    rq_activate_all_grippers(True)
    # end: URCap Program Node
  end
  $ 63 "zero_ftsensor()"
  zero_ftsensor()
  $ 64 "EXTT"
  $ 65 "Set GRP_3F_Enable=Off"
  set_standard_digital_out(4, False)
  $ 66 "Set BarcodeTrigger=Off"
  set_standard_digital_out(6, False)
  $ 67 "Set GRP_3F_Decap=Off"
  set_standard_digital_out(3, False)
  $ 68 "Set GRP_3F_Cap=Off"
  set_standard_digital_out(2, False)
  $ 69 "Set GRP_3F_Open=Off"
  set_standard_digital_out(5, False)
  $ 70 "PSE_T≔get_tool_free_pose(dir=[0,0,0.150], move_in_base_frame=True)"
  global PSE_T=get_tool_free_pose(dir=[0,0,0.150], move_in_base_frame=True)
  $ 71 "If is_reachable(Base_const, [PSE_T])"
  if (is_reachable(p[0.0,0.0,0.0,0.0,0.0,0.0], [PSE_T])):
    $ 72 "MoveL"
    $ 73 "PSE_T" "breakAfter"
    movel(PSE_T, a=1.2, v=0.15)
  end
  $ 74 "powder dispensing variable init"
  $ 75 "Start_thread≔ False "
  global Start_thread=  False
  $ 76 "vib_thread≔ False "
  global vib_thread=  False
  $ 77 "kp≔0.001"
  global kp=0.001
  $ 78 "ki≔0.00006"
  global ki=0.00006
  $ 79 "kd≔0.015"
  global kd=0.015
  $ 80 "dt≔0.03"
  global dt=0.03
  $ 81 "Integral_error≔0"
  global Integral_error=0
  $ 82 "current_error≔0"
  global current_error=0
  $ 83 "previous_error≔0"
  global previous_error=0
  $ 84 "tilt_increment≔0"
  global tilt_increment=0
  $ 85 "tilt_angle≔0"
  global tilt_angle=0
  $ 86 "diff≔0"
  global diff=0
  $ 87 "current_pose≔get_actual_tcp_pose()"
  global current_pose= get_actual_tcp_pose ()
  $ 88 "Relative_trans≔p[0, 0, -0.035, 0, 0, 0]"
  global Relative_trans=p[0, 0, -0.035, 0, 0, 0]
  $ 89 "ContA_plc_offst≔p[-0.00205, 0.02547, 0.03730, -0.03, -2.183, 6.165]"
  global ContA_plc_offst=p[-0.00205, 0.02547, 0.03730, -0.03, -2.183, 6.165]
  $ 90 "PowA_50_offset≔p[0.21808, -0.19943, 0.06584, 0, 0, 0]"
  global PowA_50_offset=p[0.21808, -0.19943, 0.06584, 0, 0, 0]
  $ 92 "tilt_init_reference()"
  tilt_init_reference()
  $ 93 "switch_spat_M≔ True "
  global switch_spat_M=  True
  $ 94 "switch_spat_S≔ True "
  global switch_spat_S=  True
  $ 95 "switch_spat_F_M≔ True "
  global switch_spat_F_M=  True
  $ 96 "switch_spat_F_S≔ True "
  global switch_spat_F_S=  True
  $ 97 "last_scale≔0"
  global last_scale=0
  $ 98 "W_EMPTY≔51.3"
  global W_EMPTY=51.3
  $ 99 "w_dosed_total≔0"
  global w_dosed_total=0
  $ 794 "Thread_1"
  thread Thread_1():
    while (True):
      $ 795 "If Start_thread≟ True "
      if (Start_thread ==   True  ):
        $ 796 "weight_value≔get_weight()"
        global weight_value=get_weight()
        $ 797 "Wait: 0.1"
        sleep(0.1)
        $ 798 "sync()"
        sync()
      end
      $ 799 "sync()"
      sync()
    end
  end
  threadId_Thread_1 = run Thread_1()
  $ 800 "Thread_2"
  thread Thread_2():
    while (True):
      $ 801 "Loop vib_thread≟ True "
      thread Thread_while_801():
        while (True):
          $ 802 "diff≔target_weight-weight_value"
          global diff=target_weight-weight_value
          $ 803 "If diff>0.02 and spatula≠'spatula_flat_S'"
          global thread_flag_803=0
          thread Thread_if_803():
            $ 805 "Set AO[0]=4.0"
            set_standard_analog_out(0, 0.4)
            thread_flag_803 = 1
          end
          if (diff>0.02  and  spatula != "spatula_flat_S"):
            global thread_handler_803=run Thread_if_803()
            while (thread_flag_803 == 0):
              if not(diff>0.02  and  spatula != "spatula_flat_S"):
                kill thread_handler_803
                thread_flag_803 = 2
              else:
                sync()
              end
            end
          else:
            thread_flag_803 = 2
          end
          if (thread_flag_803 == 2):
            $ 806 "ElseIf diff>0.02 and spatula≟'spatula_flat_S'"
            if (diff>0.02 and spatula == "spatula_flat_S"):
              $ 807 "vibration_3()"
              vibration_3()
            else:
              $ 808 "ElseIf diff≤0.03"
              global thread_flag_808=0
              thread Thread_if_808():
                $ 809 "vibration_2()"
                vibration_2()
                thread_flag_808 = 1
              end
              if (diff <= 0.03):
                global thread_handler_808=run Thread_if_808()
                while (thread_flag_808 == 0):
                  if not(diff <= 0.03):
                    kill thread_handler_808
                    thread_flag_808 = 2
                  else:
                    sync()
                  end
                end
              else:
                thread_flag_808 = 2
              end
              if (thread_flag_808 == 2):
                $ 814 "Else" "noBreak"
                $ 815 "Set AO[0]=0.0"
                set_standard_analog_out(0, 0.0)
              end
            end
          end
        end
      end
      if (vib_thread ==   True  ):
        global thread_handler_801=run Thread_while_801()
        while (vib_thread ==   True  ):
          sync()
        end
        kill thread_handler_801
      end
      $ 816 "sync()"
      sync()
    end
  end
  threadId_Thread_2 = run Thread_2()
  while (True):
    $ 100 "Robot Program"
    $ 101 "MAIN"
    $ 102 "command_manager(external_control='uGO', cond_suspend=(ITM_Manipulated and AMR_AtTarget and AMR_Charging and AMR_Battery<40), cond_unsuspend=(AMR_Battery≟60))"
    command_manager(external_control="uGO", cond_suspend=(ITM_Manipulated  and  AMR_AtTarget  and  AMR_Charging  and  AMR_Battery<40), cond_unsuspend=(AMR_Battery == 60))
    $ 103 "log_state(STATE_Info)"
    log_state(STATE_Info)
    $ 104 "Switch STATE"
    switch_1 = STATE
    $ 105 "Case 1"
    if (1 == switch_1):
      $ 106 "Stopping"
      $ 107 "STATE_Info≔'Stopping'"
      global STATE_Info="Stopping"
      $ 108 "end_freedrive_mode()"
      end_freedrive_mode()
      $ 109 "Set"
      set_tcp(p[0.0,0.0,0.161,3.1415,0.0,0.0])
      $ 110 "PSE_T≔get_tool_free_pose(dir=[0,0,0.150], move_in_base_frame=True)"
      global PSE_T=get_tool_free_pose(dir=[0,0,0.150], move_in_base_frame=True)
      $ 111 "If is_reachable(Base_const, [PSE_T])"
      if (is_reachable(p[0.0,0.0,0.0,0.0,0.0,0.0], [PSE_T])):
        $ 112 "MoveL"
        $ 113 "PSE_T" "breakAfter"
        movel(PSE_T, a=1.2, v=0.15)
      end
      $ 114 "do_transition(keep_rxry=OBJ_Picked, r=0)"
      do_transition(keep_rxry=OBJ_Picked, r=0)
      $ 123 "Call Sub_AMR_MiR_V3"
      Sub_AMR_MiR_V3()
      $ 124 "If stopping() and AMR_Done"
      if (stopping()  and  AMR_Done):
        $ 125 "STATE≔2"
        global STATE=2
        $ 126 "ugo_update_outputs()"
        ugo_update_outputs()
      end
    elif (2 == switch_1):
      $ 127 "Case 2"
      $ 128 "Stopped"
      $ 129 "STATE_Info≔'Stopped'"
      global STATE_Info="Stopped"
      $ 130 "Call Sub_AMR_MiR_V3"
      Sub_AMR_MiR_V3()
      $ 131 "If CMD_Reset  or PB_Start"
      if (CMD_Reset   or  get_standard_digital_in(0)):
        $ 132 "STATE≔3"
        global STATE=3
        $ 133 "ugo_update_outputs()"
        ugo_update_outputs()
      end
    elif (3 == switch_1):
      $ 134 "Case 3"
      $ 135 " Resetting"
      $ 136 "STATE_Info≔'Resetting'"
      global STATE_Info="Resetting"
      $ 137 "uML"
      $ 138 "reset_error()"
      reset_error()
      $ 139 "reset_warning()"
      reset_warning()
      $ 140 "PROCESS_Step≔0"
      global PROCESS_Step=0
      $ 141 "PROCESS_Info≔''"
      global PROCESS_Info=""
      $ 142 "ARM_Referenced≔ False "
      global ARM_Referenced=  False
      $ 143 "WRK_Done≔ False "
      global WRK_Done=  False
      $ 144 "ITM_Prepared≔ False "
      global ITM_Prepared=  False
      $ 145 "ITM_Manipulated≔ False "
      global ITM_Manipulated=  False
      $ 146 "STP≔0"
      global STP=0
      $ 147 "Action≔0"
      global Action=0
      $ 148 "Action_Info≔''"
      global Action_Info=""
      $ 149 "ITM_ID≔0"
      global ITM_ID=0
      $ 150 "JIG≔0"
      global JIG=0
      $ 151 "JIG_Slot≔0"
      global JIG_Slot=0
      $ 152 "Task_info≔''"
      global Task_info=""
      $ 153 "Set"
      set_tcp(p[0.0,0.0,0.161,3.1415,0.0,0.0])
      $ 154 "App"
      $ 155 "'ADD APPLICATION SPECIFIC COMMANDS'"
      # 'ADD APPLICATION SPECIFIC COMMANDS'
      $ 156 "OBJ_Type≔0"
      global OBJ_Type=0
      $ 157 "OBJ_Nbr≔0"
      global OBJ_Nbr=0
      $ 158 "If CNT_Rack_Output≥50"
      if (CNT_Rack_Output >= 50):
        $ 159 "CNT_Rack_Output≔0"
        global CNT_Rack_Output=0
      end
      $ 160 "TASK≔struct(ID=0, NAVI=struct(target=0, footprint=0, protectiveOff=0, dock=0), WORK=struct(ITM_ID_Src=0, JIG_ID_Src=0, OBJ_Nbr_Src=0, ACT_Src=0, ITM_ID_Tgt=0, JIG_ID_Tgt=0, OBJ_Nbr_Tgt=0, ACT_Tgt=0, OBJ_Type=0))"
      global TASK=struct(ID=0, NAVI=struct(target=0, footprint=0, protectiveOff=0, dock=0), WORK=struct(ITM_ID_Src=0, JIG_ID_Src=0, OBJ_Nbr_Src=0, ACT_Src=0, ITM_ID_Tgt=0, JIG_ID_Tgt=0, OBJ_Nbr_Tgt=0, ACT_Tgt=0, OBJ_Type=0))
      $ 161 "Call Sub_AMR_MiR_V3"
      Sub_AMR_MiR_V3()
      $ 162 "If resetting() and AMR_Done"
      if (resetting()  and  AMR_Done):
        $ 163 "STATE≔4"
        global STATE=4
        $ 164 "ugo_update_outputs()"
        ugo_update_outputs()
      end
    elif (4 == switch_1):
      $ 165 "Case 4"
      $ 166 "Idle"
      $ 167 "STATE_Info≔'Idle'"
      global STATE_Info="Idle"
      $ 168 "If CMD_Start"
      if (CMD_Start):
        $ 169 "STATE≔5"
        global STATE=5
        $ 170 "ugo_update_outputs()"
        ugo_update_outputs()
      end
    elif (5 == switch_1):
      $ 171 "Case 5"
      $ 172 "Starting"
      $ 173 "STATE_Info≔'Starting'"
      global STATE_Info="Starting"
      $ 174 "'ADD COMMANDS WHAT TO START WITH'"
      # 'ADD COMMANDS WHAT TO START WITH'
      $ 175 "Call Sub_AMR_MiR_V3"
      Sub_AMR_MiR_V3()
      $ 176 "get ugo data"
      $ 177 "Assign Tasks"
      $ 178 "TASK.ID = ugo_get_task()"
      TASK.ID = ugo_get_task()
      $ 179 "If TASK.ID≟1"
      if (TASK.ID == 1):
        $ 180 "Task_info≔'Charge'"
        global Task_info="Charge"
        $ 181 "Parameters"
        $ 182 "AMR_PosTarget≔1"
        global AMR_PosTarget=1
      else:
        $ 183 "ElseIf TASK.ID≟9"
        if (TASK.ID == 9):
          $ 184 "'Pick Sarstedt Rack from Variable source'"
          # 'Pick Sarstedt Rack from Variable source'
          $ 185 "Task_info≔'Navigate to Target'"
          global Task_info="Navigate to Target"
          $ 186 "Parameters"
          $ 187 "AMR_PosTarget≔UGO.read_input('00','ITM_ID')"
          global AMR_PosTarget=UGO.read_input("00","ITM_ID")
        else:
          $ 188 "ElseIf TASK.ID≟49"
          if (TASK.ID == 49):
            $ 189 "Task_info≔'Pick Containers'"
            global Task_info="Pick Containers"
            $ 190 "Parameters"
            $ 191 "ITM_ID≔1"
            global ITM_ID=1
            $ 192 "OBJ_Type≔6"
            global OBJ_Type=6
            $ 193 "JIG≔15"
            global JIG=15
            $ 194 "AMR_PosTarget≔3"
            global AMR_PosTarget=3
          else:
            $ 195 "ElseIf TASK.ID≟50"
            if (TASK.ID == 50):
              $ 196 "Task_info≔'Decap Containers'"
              global Task_info="Decap Containers"
              $ 197 "Parameters"
              $ 198 "ITM_ID≔1"
              global ITM_ID=1
              $ 199 "OBJ_Type≔6"
              global OBJ_Type=6
              $ 200 "JIG≔16"
              global JIG=16
              $ 201 "AMR_PosTarget≔5"
              global AMR_PosTarget=5
            else:
              $ 202 "ElseIf TASK.ID≟51"
              if (TASK.ID == 51):
                $ 203 "Task_info≔'Detect Spatula and transfer powder'"
                global Task_info="Detect Spatula and transfer powder"
                $ 204 "Parameters"
                $ 205 "ITM_ID≔1"
                global ITM_ID=1
                $ 206 "target_weight≔(UGO.read_input('00','Target_weight'))/1000"
                global target_weight=(UGO.read_input("00","Target_weight"))/1000
                $ 207 "OBJ_Type≔8"
                global OBJ_Type=8
                $ 208 "JIG≔16"
                global JIG=16
                $ 209 "AMR_PosTarget≔5"
                global AMR_PosTarget=5
              else:
                $ 210 "ElseIf TASK.ID≟52"
                if (TASK.ID == 52):
                  $ 211 "Task_info≔'Pick Powder'"
                  global Task_info="Pick Powder"
                  $ 212 "Parameters"
                  $ 213 "ITM_ID≔1"
                  global ITM_ID=1
                  $ 214 "OBJ_Type≔6"
                  global OBJ_Type=6
                  $ 215 "JIG≔15"
                  global JIG=15
                  $ 216 "AMR_PosTarget≔3"
                  global AMR_PosTarget=3
                else:
                  $ 217 "ElseIf TASK.ID≟53"
                  if (TASK.ID == 53):
                    $ 218 "Task_info≔'Decap Powder'"
                    global Task_info="Decap Powder"
                    $ 219 "Parameters"
                    $ 220 "ITM_ID≔1"
                    global ITM_ID=1
                    $ 221 "OBJ_Type≔6"
                    global OBJ_Type=6
                    $ 222 "JIG≔1"
                    global JIG=1
                    $ 223 "AMR_PosTarget≔5"
                    global AMR_PosTarget=5
                  else:
                    $ 224 "ElseIf TASK.ID≟54"
                    if (TASK.ID == 54):
                      $ 225 "Task_info≔'Empty and swap Powder container'"
                      global Task_info="Empty and swap Powder container"
                      $ 234 "Parameters"
                      $ 235 "ITM_ID≔1"
                      global ITM_ID=1
                      $ 237 "W_now≔(UGO.read_input('00','Container_weight'))/1000"
                      global W_now=(UGO.read_input("00","Container_weight"))/1000
                      $ 238 "Pow_name≔(UGO.read_input('00','Powder_name'))"
                      global Pow_name=(UGO.read_input("00","Powder_name"))
                      $ 239 "scooping_init()"
                      scooping_init()
                      $ 240 "target_weight≔W_now-W_EMPTY-(0.002*W_FULL)"
                      global target_weight=W_now-W_EMPTY-(0.002*W_FULL)
                      $ 241 "OBJ_Type≔6"
                      global OBJ_Type=6
                      $ 242 "JIG≔17"
                      global JIG=17
                      $ 243 "AMR_PosTarget≔5"
                      global AMR_PosTarget=5
                    else:
                      $ 244 "ElseIf TASK.ID≟55"
                      if (TASK.ID == 55):
                        $ 245 "Task_info≔'Place Powder'"
                        global Task_info="Place Powder"
                        $ 246 "Parameters"
                        $ 247 "ITM_ID≔1"
                        global ITM_ID=1
                        $ 248 "OBJ_Type≔6"
                        global OBJ_Type=6
                        $ 249 "JIG≔21"
                        global JIG=21
                        $ 250 "AMR_PosTarget≔5"
                        global AMR_PosTarget=5
                      else:
                        $ 251 "ElseIf TASK.ID≟56"
                        if (TASK.ID == 56):
                          $ 252 "Task_info≔'Dose Powder'"
                          global Task_info="Dose Powder"
                          $ 253 "Parameters"
                          $ 254 "ITM_ID≔1"
                          global ITM_ID=1
                          $ 255 "target_weight≔(UGO.read_input('00','Target_weight'))/1000"
                          global target_weight=(UGO.read_input("00","Target_weight"))/1000
                          $ 256 "W_now≔(UGO.read_input('00','Container_weight'))/1000"
                          global W_now=(UGO.read_input("00","Container_weight"))/1000
                          $ 258 "Pow_name≔(UGO.read_input('00','Powder_name'))"
                          global Pow_name=(UGO.read_input("00","Powder_name"))
                          $ 259 "OBJ_Type≔6"
                          global OBJ_Type=6
                          $ 260 "JIG≔17"
                          global JIG=17
                          $ 261 "AMR_PosTarget≔5"
                          global AMR_PosTarget=5
                        else:
                          $ 262 "ElseIf TASK.ID≟57"
                          if (TASK.ID == 57):
                            $ 263 "Task_info≔'Recipe Powder dosing'"
                            global Task_info="Recipe Powder dosing"
                            $ 264 "Parameters"
                            $ 265 "ITM_ID≔1"
                            global ITM_ID=1
                            $ 266 "Pow_A≔(UGO.read_input('00','PowderA'))"
                            global Pow_A=(UGO.read_input("00","PowderA"))
                            $ 267 "Pow_B≔(UGO.read_input('00','PowderB'))"
                            global Pow_B=(UGO.read_input("00","PowderB"))
                            $ 268 "Pow_C≔(UGO.read_input('00','PowderC'))"
                            global Pow_C=(UGO.read_input("00","PowderC"))
                            $ 269 "Total_weight≔(UGO.read_input('00','Total_weight'))/1000"
                            global Total_weight=(UGO.read_input("00","Total_weight"))/1000
                            $ 270 "Pow_A_percent≔(UGO.read_input('00','PowderA_percentage'))/100"
                            global Pow_A_percent=(UGO.read_input("00","PowderA_percentage"))/100
                            $ 271 "Pow_B_percent≔(UGO.read_input('00','PowderB_percentage'))/100"
                            global Pow_B_percent=(UGO.read_input("00","PowderB_percentage"))/100
                            $ 272 "Pow_C_percent≔(UGO.read_input('00','PowderC_percentage'))/100"
                            global Pow_C_percent=(UGO.read_input("00","PowderC_percentage"))/100
                            $ 273 "OBJ_Type≔6"
                            global OBJ_Type=6
                            $ 274 "JIG≔17"
                            global JIG=17
                            $ 275 "AMR_PosTarget≔5"
                            global AMR_PosTarget=5
                          else:
                            $ 276 "ElseIf TASK.ID≟58"
                            if (TASK.ID == 58):
                              $ 277 "Task_info≔'Pick Powder containers'"
                              global Task_info="Pick Powder containers"
                              $ 278 "Parameters"
                              $ 279 "ITM_ID≔1"
                              global ITM_ID=1
                              $ 280 "OBJ_Type≔6"
                              global OBJ_Type=6
                              $ 281 "JIG≔15"
                              global JIG=15
                              $ 282 "AMR_PosTarget≔3"
                              global AMR_PosTarget=3
                            else:
                              $ 283 "ElseIf TASK.ID≟59"
                              if (TASK.ID == 59):
                                $ 284 "Task_info≔'Calibration for new powder'"
                                global Task_info="Calibration for new powder"
                                $ 285 "Parameters"
                                $ 286 "ITM_ID≔1"
                                global ITM_ID=1
                                $ 287 "Pow_name≔(UGO.read_input('00','Pow_name'))"
                                global Pow_name=(UGO.read_input("00","Pow_name"))
                                $ 288 "W_now≔(UGO.read_input('00','Container_weight'))/1000"
                                global W_now=(UGO.read_input("00","Container_weight"))/1000
                                $ 289 "density≔(UGO.read_input('00', 'Density'))"
                                global density=(UGO.read_input("00", "Density"))
                                $ 290 "Flowability≔(UGO.read_input('00', 'Flowability'))"
                                global Flowability=(UGO.read_input("00", "Flowability"))
                                $ 291 "spatula≔(UGO.read_input('00','Spatula'))"
                                global spatula=(UGO.read_input("00","Spatula"))
                                $ 292 "OBJ_Type≔6"
                                global OBJ_Type=6
                                $ 293 "JIG≔17"
                                global JIG=17
                                $ 294 "AMR_PosTarget≔5"
                                global AMR_PosTarget=5
                              else:
                                $ 295 "Else" "noBreak"
                                $ 296 "set_error(ERROR_WRONG_ORDER)"
                                set_error(ERROR_WRONG_ORDER)
                              end
                            end
                          end
                        end
                      end
                    end
                  end
                end
              end
            end
          end
        end
      end
      $ 297 "test ugo"
      $ 298 "Wait: 0.2"
      sleep(0.2)
      $ 299 "ugo_update_outputs()"
      ugo_update_outputs()
      $ 300 "If starting() and AMR_Done"
      if (starting()  and  AMR_Done):
        $ 301 "log_message(Task_info, 'New Task: ')"
        log_message(Task_info, "New Task: ")
        $ 302 "log_message(to_str(TASK.ID), 'Task_ID: ')"
        log_message(to_str(TASK.ID), "Task_ID: ")
        $ 303 "do_transition(keep_rxry=OBJ_Picked)"
        do_transition(keep_rxry=OBJ_Picked)
        $ 304 "STATE≔6"
        global STATE=6
        $ 305 "ugo_update_outputs()"
        ugo_update_outputs()
      end
    elif (6 == switch_1):
      $ 306 "Case 6"
      $ 307 "Execute"
      $ 308 "STATE_Info≔'Execute'"
      global STATE_Info="Execute"
      $ 309 "If  not CMD_Hold and not CMD_Suspend"
      global thread_flag_309=0
      thread Thread_if_309():
        $ 310 "Switch PROCESS_Step"
        switch_2 = PROCESS_Step
        $ 311 "Case 0"
        if (0 == switch_2):
          $ 312 "PROCESS_Info≔'process control'"
          global PROCESS_Info="process control"
          $ 313 "log_process(PROCESS_Info)"
          log_process(PROCESS_Info)
          $ 314 "process control"
          $ 315 "If  not AMR_AtTarget"
          if (  not  AMR_AtTarget):
            $ 316 "PROCESS_Step≔1"
            global PROCESS_Step=1
          else:
            $ 317 "ElseIf (( not ITM_Prepared and  not WRK_Done) or (ITM_Prepared and WRK_Done))"
            if (((  not  ITM_Prepared  and    not  WRK_Done)  or  (ITM_Prepared  and  WRK_Done))):
              $ 318 "PROCESS_Step≔2"
              global PROCESS_Step=2
            else:
              $ 319 "ElseIf  not WRK_Done"
              if (  not  WRK_Done):
                $ 320 "PROCESS_Step≔3"
                global PROCESS_Step=3
              else:
                $ 321 "Else" "noBreak"
                $ 322 "task finished"
                $ 323 "PROCESS_Info≔''"
                global PROCESS_Info=""
                $ 324 "STATE≔7"
                global STATE=7
                $ 325 "ugo_update_outputs()"
                ugo_update_outputs()
              end
            end
          end
        elif (1 == switch_2):
          $ 326 "Case 1"
          $ 327 "navigate"
          $ 328 "'MOVING THE uML'"
          # 'MOVING THE uML'
          $ 329 "PROCESS_Info≔'move to target'"
          global PROCESS_Info="move to target"
          $ 330 "log_process(PROCESS_Info)"
          log_process(PROCESS_Info)
          $ 331 "If TASK.ID≟1"
          if (TASK.ID == 1):
            $ 332 "Action≔51"
            global Action=51
          else:
            $ 333 "Else" "noBreak"
            $ 334 "Action≔52"
            global Action=52
          end
          $ 335 "Call Sub_AMR_MiR_V3"
          Sub_AMR_MiR_V3()
          $ 336 "If AMR_Done"
          if (AMR_Done):
            $ 337 "PROCESS_Step≔0"
            global PROCESS_Step=0
          end
        elif (2 == switch_2):
          $ 338 "Case 2"
          $ 339 "prepare"
          $ 340 "'THINGS THAT HAVE TO BE DONE ONCE IN A SEQUENCE,WORKFLOW'"
          # 'THINGS THAT HAVE TO BE DONE ONCE IN A SEQUENCE,WORKFLOW'
          $ 341 "PROCESS_Info≔'prepare for work'"
          global PROCESS_Info="prepare for work"
          $ 342 "log_process(PROCESS_Info)"
          log_process(PROCESS_Info)
          $ 343 "If TASK.WORK.ITM_ID_Src>1"
          if (TASK.WORK.ITM_ID_Src>1):
            $ 344 "ITM_ID≔TASK.WORK.ITM_ID_Src"
            global ITM_ID=TASK.WORK.ITM_ID_Src
          else:
            $ 345 "ElseIf TASK.WORK.ITM_ID_Tgt>1"
            if (TASK.WORK.ITM_ID_Tgt>1):
              $ 346 "ITM_ID≔TASK.WORK.ITM_ID_Tgt"
              global ITM_ID=TASK.WORK.ITM_ID_Tgt
            end
          end
          $ 347 "If  not ARM_Referenced and (ITM_ID≠0)"
          if (  not  ARM_Referenced  and  (ITM_ID != 0)):
            $ 348 "STP≔1"
            global STP=1
          else:
            $ 349 "ElseIf ARM_Referenced or (ITM_ID≟0)"
            if (ARM_Referenced  or  (ITM_ID == 0)):
              $ 350 "STP≔2"
              global STP=2
            end
          end
          $ 351 "Switch STP"
          switch_3 = STP
          $ 352 "Case 1"
          if (1 == switch_3):
            $ 353 "reference"
            $ 354 "STP_Info≔'reference at target position'"
            global STP_Info="reference at target position"
            $ 355 "log_step(STP_Info)"
            log_step(STP_Info)
            $ 356 "If ITM_ID≟1"
            if (ITM_ID == 1):
              $ 357 "CAM_Done≔ True "
              global CAM_Done=  True
            else:
              $ 358 "Else" "noBreak"
              $ 359 "Action≔131"
              global Action=131
              $ 360 "Call Sub_Vision_V18"
              Sub_Vision_V18()
            end
            $ 362 "If CAM_Done and  not ERROR.FLAG"
            if (CAM_Done  and    not  ERROR.FLAG):
              $ 363 "log_step('ARM referenced')"
              log_step("ARM referenced")
              $ 364 "ARM_Referenced≔ True "
              global ARM_Referenced=  True
            end
          elif (2 == switch_3):
            $ 365 "Case 2"
            $ 366 "manipulate"
            $ 367 "STP_Info≔'manipulate item'"
            global STP_Info="manipulate item"
            $ 368 "log_step(STP_Info)"
            log_step(STP_Info)
            $ 369 "'In case pressing button is needed'"
            # 'In case pressing button is needed'
            $ 370 "If found_in_list(ITM_ID, ITM_ID_List)"
            if (found_in_list(ITM_ID, ITM_ID_List)):
              $ 371 "Switch ITM_ID"
              switch_4 = ITM_ID
              $ 372 "Case 0"
              if (0 == switch_4):
                $ 373 "ITM_Manipulated≔ not ITM_Manipulated"
                global ITM_Manipulated=  not  ITM_Manipulated
              elif (1 == switch_4):
                $ 374 "Case 1"
                $ 375 "ITM_Manipulated≔ not ITM_Manipulated"
                global ITM_Manipulated=  not  ITM_Manipulated
              elif (2 == switch_4):
                $ 376 "Case 2"
              else:
                $ 386 "Default Case"
                $ 387 "ITM_Manipulated≔ not ITM_Manipulated"
                global ITM_Manipulated=  not  ITM_Manipulated
              end
            end
          end
          $ 388 "ITM_Prepared≔(ITM_Manipulated or  not found_in_list(ITM_ID, ITM_ID_List)) and (ARM_Referenced or ITM_ID≟0) and  not WRK_Done"
          global ITM_Prepared=(ITM_Manipulated  or    not  found_in_list(ITM_ID, ITM_ID_List))  and  (ARM_Referenced  or  ITM_ID == 0)  and    not  WRK_Done
          $ 389 "STP≔0"
          global STP=0
          $ 390 "STP_Info≔''"
          global STP_Info=""
          $ 391 "PROCESS_Step≔0"
          global PROCESS_Step=0
        elif (3 == switch_2):
          $ 392 "Case 3"
          $ 393 "work"
          $ 394 "'ADD EVERY MACHINE, OBJECT, STATION TO WORK ON'"
          # 'ADD EVERY MACHINE, OBJECT, STATION TO WORK ON'
          $ 395 "Switch ITM_ID"
          switch_3 = ITM_ID
          $ 396 "Case 1"
          if (1 == switch_3):
            $ 397 "uLM"
            $ 398 "If TASK.ID≟12"
            if (TASK.ID == 12):
              $ 399 "fill racks"
              $ 400 "Action≔151"
              global Action=151
              $ 401 "Call Sub_Vision_V18"
              Sub_Vision_V18()
              $ 402 "If  not ERROR.FLAG"
              if (  not  ERROR.FLAG):
                $ 403 "Actions for the task"
                $ 404 "Action≔1"
                global Action=1
                $ 405 "JIG≔2"
                global JIG=2
                $ 406 "JIG_Slot≔CAM_Result[0]"
                global JIG_Slot=CAM_Result[0]
                $ 407 "OBJ_Nbr≔CAM_Result[0]"
                global OBJ_Nbr=CAM_Result[0]
                $ 408 "OBJ_Type≔2"
                global OBJ_Type=2
                $ 409 "Call Sub_Action_V4"
                Sub_Action_V4()
                $ 410 "If OBJ_Picked"
                if (OBJ_Picked):
                  $ 411 "CAM_Result.remove(0)"
                  CAM_Result.remove(0)
                  $ 412 "PRC_TubCounter≔PRC_TubCounter+1"
                  global PRC_TubCounter=PRC_TubCounter+1
                  $ 413 "If PRC_TubCounter%4≟0"
                  if (PRC_TubCounter%4 == 0):
                    $ 414 "JIG_Slot≔4"
                    global JIG_Slot=4
                  else:
                    $ 415 "Else" "noBreak"
                    $ 416 "JIG_Slot≔PRC_TubCounter%4"
                    global JIG_Slot=PRC_TubCounter%4
                  end
                  $ 417 "OBJ_Nbr≔ceil(PRC_TubCounter/4)"
                  global OBJ_Nbr=ceil(PRC_TubCounter/4)
                  $ 418 "Action≔2"
                  global Action=2
                  $ 419 "JIG≔4"
                  global JIG=4
                  $ 420 "Call Sub_Action_V4"
                  Sub_Action_V4()
                  $ 421 "Action≔151"
                  global Action=151
                  $ 422 "Call Sub_Vision_V18"
                  Sub_Vision_V18()
                end
              end
              $ 423 "If (CAM_Captures≥CAM_PRM_Retries) or (PRC_TubCounter≥32)"
              if ((CAM_Captures >= CAM_PRM_Retries)  or  (PRC_TubCounter >= 32)):
                $ 424 "PROCESS_Step≔0"
                global PROCESS_Step=0
                $ 425 "WRK_Done≔ True "
                global WRK_Done=  True
              end
            else:
              $ 426 "ElseIf TASK.ID≟49"
              if (TASK.ID == 49):
                $ 427 "Pick Powder container"
                $ 428 "Action≔131"
                global Action=131
                $ 429 "Call Sub_Vision_V18"
                Sub_Vision_V18()
                $ 430 "Action≔35"
                global Action=35
                $ 431 "Call Sub_Action_V4"
                Sub_Action_V4()
                $ 432 "PROCESS_Step≔0"
                global PROCESS_Step=0
                $ 433 "WRK_Done≔ True "
                global WRK_Done=  True
              else:
                $ 434 "ElseIf TASK.ID≟50"
                if (TASK.ID == 50):
                  $ 435 "Decap containers"
                  $ 436 "Action≔36"
                  global Action=36
                  $ 437 "Call Sub_Action_V4"
                  Sub_Action_V4()
                  $ 438 "PROCESS_Step≔0"
                  global PROCESS_Step=0
                  $ 439 "WRK_Done≔ True "
                  global WRK_Done=  True
                else:
                  $ 440 "ElseIf TASK.ID≟51"
                  if (TASK.ID == 51):
                    $ 441 "Detect Spatula and transfer powder"
                    $ 442 "Action≔131"
                    global Action=131
                    $ 443 "Call Sub_Vision_V18"
                    Sub_Vision_V18()
                    $ 444 "Action≔37"
                    global Action=37
                    $ 445 "Call Sub_Action_V4"
                    Sub_Action_V4()
                    $ 446 "PROCESS_Step≔0"
                    global PROCESS_Step=0
                    $ 447 "WRK_Done≔ True "
                    global WRK_Done=  True
                  else:
                    $ 448 "ElseIf TASK.ID≟52"
                    if (TASK.ID == 52):
                      $ 449 "Pick Powder container"
                      $ 450 "Action≔131"
                      global Action=131
                      $ 451 "Call Sub_Vision_V18"
                      Sub_Vision_V18()
                      $ 452 "Action≔39"
                      global Action=39
                      $ 453 "Call Sub_Action_V4"
                      Sub_Action_V4()
                      $ 454 "PROCESS_Step≔0"
                      global PROCESS_Step=0
                      $ 455 "WRK_Done≔ True "
                      global WRK_Done=  True
                    else:
                      $ 456 "ElseIf TASK.ID≟53"
                      if (TASK.ID == 53):
                        $ 457 "Decap containerA"
                        $ 458 "Action≔40"
                        global Action=40
                        $ 459 "Call Sub_Action_V4"
                        Sub_Action_V4()
                        $ 460 "PROCESS_Step≔0"
                        global PROCESS_Step=0
                        $ 461 "WRK_Done≔ True "
                        global WRK_Done=  True
                      else:
                        $ 462 "ElseIf TASK.ID≟55"
                        if (TASK.ID == 55):
                          $ 463 "Place Powder"
                          $ 464 "Action≔131"
                          global Action=131
                          $ 465 "Call Sub_Vision_V18"
                          Sub_Vision_V18()
                          $ 466 "Action≔41"
                          global Action=41
                          $ 467 "Call Sub_Action_V4"
                          Sub_Action_V4()
                          $ 468 "PROCESS_Step≔0"
                          global PROCESS_Step=0
                          $ 469 "WRK_Done≔ True "
                          global WRK_Done=  True
                        else:
                          $ 470 "ElseIf TASK.ID≟54"
                          if (TASK.ID == 54):
                            $ 471 "Empty and swap container"
                            $ 472 "Action≔131"
                            global Action=131
                            $ 473 "Call Sub_Vision_V18"
                            Sub_Vision_V18()
                            $ 474 "Action≔42"
                            global Action=42
                            $ 475 "Call Sub_Action_V4"
                            Sub_Action_V4()
                            $ 476 "PROCESS_Step≔0"
                            global PROCESS_Step=0
                            $ 477 "WRK_Done≔ True "
                            global WRK_Done=  True
                          else:
                            $ 478 "ElseIf TASK.ID≟56"
                            if (TASK.ID == 56):
                              $ 479 "Dispense Powder"
                              $ 480 "Action≔131"
                              global Action=131
                              $ 481 "Call Sub_Vision_V18"
                              Sub_Vision_V18()
                              $ 482 "Action≔43"
                              global Action=43
                              $ 483 "Call Sub_Action_V4"
                              Sub_Action_V4()
                              $ 484 "PROCESS_Step≔0"
                              global PROCESS_Step=0
                              $ 485 "WRK_Done≔ True "
                              global WRK_Done=  True
                            else:
                              $ 486 "ElseIf TASK.ID≟57"
                              if (TASK.ID == 57):
                                $ 487 "Recipe Dosing"
                                $ 488 "QR_Action≔1"
                                global QR_Action=1
                                $ 489 "Action≔48"
                                global Action=48
                                $ 490 "Call Sub_Action_V4"
                                Sub_Action_V4()
                                $ 491 "recipe_init(Pow_A, Pow_B, Pow_C, Total_weight, Pow_A_percent, Pow_B_percent, Pow_C_percent)"
                                recipe_init(Pow_A, Pow_B, Pow_C, Total_weight, Pow_A_percent, Pow_B_percent, Pow_C_percent)
                                $ 492 "Loop recipe_next()≟ True "
                                while (recipe_next() ==   True  ):
                                  $ 493 "Action≔44"
                                  global Action=44
                                  $ 494 "Call Sub_Action_V4"
                                  Sub_Action_V4()
                                  $ 495 "JIG≔21"
                                  global JIG=21
                                  $ 496 "Action≔131"
                                  global Action=131
                                  $ 497 "Call Sub_Vision_V18"
                                  Sub_Vision_V18()
                                  $ 498 "Action≔45"
                                  global Action=45
                                  $ 499 "Call Sub_Action_V4"
                                  Sub_Action_V4()
                                  $ 500 "dosing_start()"
                                  dosing_start()
                                  $ 501 "JIG≔17"
                                  global JIG=17
                                  $ 502 "Action≔131"
                                  global Action=131
                                  $ 503 "Call Sub_Vision_V18"
                                  Sub_Vision_V18()
                                  $ 504 "Action≔46"
                                  global Action=46
                                  $ 505 "Call Sub_Action_V4"
                                  Sub_Action_V4()
                                  $ 506 "dosing_end()"
                                  dosing_end()
                                end
                                $ 507 "PROCESS_Step≔0"
                                global PROCESS_Step=0
                                $ 508 "WRK_Done≔ True "
                                global WRK_Done=  True
                              else:
                                $ 509 "ElseIf TASK.ID≟58"
                                if (TASK.ID == 58):
                                  $ 510 "Pick Powder containers"
                                  $ 511 "Num_cont_picked≔0"
                                  global Num_cont_picked=0
                                  $ 512 "powder_position≔'Position1'"
                                  global powder_position="Position1"
                                  $ 513 "Loop Num_cont_picked<3"
                                  while (Num_cont_picked<3):
                                    $ 514 "Action≔131"
                                    global Action=131
                                    $ 515 "Call Sub_Vision_V18"
                                    Sub_Vision_V18()
                                    $ 516 "Action≔47"
                                    global Action=47
                                    $ 517 "Call Sub_Action_V4"
                                    Sub_Action_V4()
                                  end
                                  $ 518 "PROCESS_Step≔0"
                                  global PROCESS_Step=0
                                  $ 519 "WRK_Done≔ True "
                                  global WRK_Done=  True
                                else:
                                  $ 520 "ElseIf TASK.ID≟59"
                                  if (TASK.ID == 59):
                                    $ 521 "Calibration"
                                    $ 525 "Action≔49"
                                    global Action=49
                                    $ 526 "Call Sub_Action_V4"
                                    Sub_Action_V4()
                                    $ 527 "PROCESS_Step≔0"
                                    global PROCESS_Step=0
                                    $ 528 "WRK_Done≔ True "
                                    global WRK_Done=  True
                                  end
                                end
                              end
                            end
                          end
                        end
                      end
                    end
                  end
                end
              end
            end
          elif (2 == switch_3):
            $ 529 "Case 2"
          elif (5 == switch_3):
            $ 571 "Case 5"
          elif (20 == switch_3):
            $ 579 "Case 20"
          elif (43 == switch_3):
            $ 641 "Case 43"
          else:
            $ 649 "Default Case"
            $ 650 "WRK_Done≔ True "
            global WRK_Done=  True
            $ 651 "PROCESS_Step≔0"
            global PROCESS_Step=0
          end
        end
        thread_flag_309 = 1
      end
      if (  not  CMD_Hold and not CMD_Suspend):
        global thread_handler_309=run Thread_if_309()
        while (thread_flag_309 == 0):
          if not(  not  CMD_Hold and not CMD_Suspend):
            kill thread_handler_309
            thread_flag_309 = 2
          else:
            sync()
          end
        end
      else:
        thread_flag_309 = 2
      end
      $ 652 "If CMD_Hold"
      if (CMD_Hold):
        $ 653 "STATE≔9"
        global STATE=9
        $ 654 "ugo_update_outputs()"
        ugo_update_outputs()
      else:
        $ 655 "ElseIf CMD_Suspend"
        if (CMD_Suspend):
          $ 656 "STATE≔12"
          global STATE=12
          $ 657 "ugo_update_outputs()"
          ugo_update_outputs()
        end
      end
    elif (7 == switch_1):
      $ 658 "Case 7"
      $ 659 "Completing"
      $ 660 "STATE_Info≔'Completing'"
      global STATE_Info="Completing"
      $ 661 "'ADD COMMANDS FOR COMPLETING THE PROCESS'"
      # 'ADD COMMANDS FOR COMPLETING THE PROCESS'
      $ 662 "do_transition(keep_rxry=OBJ_Picked)"
      do_transition(keep_rxry=OBJ_Picked)
      $ 663 "Call Sub_AMR_MiR_V3"
      Sub_AMR_MiR_V3()
      $ 664 "If completing() and AMR_Done"
      if (completing()  and  AMR_Done):
        $ 665 "STATE≔8"
        global STATE=8
        $ 666 "ugo_update_outputs()"
        ugo_update_outputs()
      end
    elif (8 == switch_1):
      $ 667 "Case 8"
      $ 668 "Complete"
      $ 669 "STATE_Info≔'Complete'"
      global STATE_Info="Complete"
      $ 670 "If CMD_Reset"
      if (CMD_Reset):
        $ 671 "STATE≔3"
        global STATE=3
        $ 672 "ugo_update_outputs()"
        ugo_update_outputs()
      end
    elif (9 == switch_1):
      $ 673 "Case 9"
      $ 674 "Holding"
      $ 675 "STATE_Info≔'Holding'"
      global STATE_Info="Holding"
      $ 676 "stopl(0.5)"
      stopl(0.5)
      $ 677 "Call Sub_AMR_MiR_V3"
      Sub_AMR_MiR_V3()
      $ 678 "If holding() and AMR_Done"
      if (holding()  and  AMR_Done):
        $ 679 "STATE≔10"
        global STATE=10
        $ 680 "ugo_update_outputs()"
        ugo_update_outputs()
      end
    elif (10 == switch_1):
      $ 681 "Case 10"
      $ 682 "Held"
      $ 683 "STATE_Info≔'Held'"
      global STATE_Info="Held"
      $ 684 "If CMD_Unhold"
      if (CMD_Unhold):
        $ 685 "end_freedrive_mode()"
        end_freedrive_mode()
        $ 686 "STATE≔11"
        global STATE=11
        $ 687 "ugo_update_outputs()"
        ugo_update_outputs()
      else:
        $ 688 "ElseIf FNC_Freedrive"
        if (FNC_Freedrive):
          $ 689 "freedrive_mode()"
          freedrive_mode()
        else:
          $ 690 "Else" "noBreak"
          $ 691 "end_freedrive_mode()"
          end_freedrive_mode()
        end
      end
    elif (11 == switch_1):
      $ 692 "Case 11"
      $ 693 "Unholding"
      $ 694 "STATE_Info≔'Unholding'"
      global STATE_Info="Unholding"
      $ 695 "Clearing"
      $ 696 "Switch ERROR.ID"
      switch_2 = ERROR.ID
      $ 697 "Case 1002"
      if (1002 == switch_2):
        $ 698 "AMR_AtTarget≔ False "
        global AMR_AtTarget=  False
        $ 699 "ARM_Referenced≔ False "
        global ARM_Referenced=  False
        $ 700 "ITM_Prepared≔ False "
        global ITM_Prepared=  False
        $ 701 "PROCESS_Step≔1"
        global PROCESS_Step=1
      elif (2007 == switch_2):
        $ 702 "Case 2007"
        $ 703 "PROCESS_Step≔1"
        global PROCESS_Step=1
      end
      $ 704 "reset_error()"
      reset_error()
      $ 705 "reset_warning()"
      reset_warning()
      $ 706 "OBJ_Picked≔gripper_has_object()"
      global OBJ_Picked=gripper_has_object()
      $ 707 "Call Sub_AMR_MiR_V3"
      Sub_AMR_MiR_V3()
      $ 708 "If unholding() and AMR_Done"
      if (unholding()  and  AMR_Done):
        $ 709 "STATE≔6"
        global STATE=6
        $ 710 "ugo_update_outputs()"
        ugo_update_outputs()
      end
    elif (12 == switch_1):
      $ 711 "Case 12"
      $ 712 "Suspending"
      $ 713 "STATE_Info≔'Suspending'"
      global STATE_Info="Suspending"
      $ 714 "PROCESS_Info≔str_cat(PROCESS_Info, ' suspended')"
      global PROCESS_Info=str_cat(PROCESS_Info, " suspended")
      $ 715 "If suspending()"
      if (suspending()):
        $ 716 "STATE≔13"
        global STATE=13
        $ 717 "ugo_update_outputs()"
        ugo_update_outputs()
      end
    elif (13 == switch_1):
      $ 718 "Case 13"
      $ 719 "Suspended"
      $ 720 "STATE_Info≔'Suspended'"
      global STATE_Info="Suspended"
      $ 721 "Call Sub_AMR_MiR_V3"
      Sub_AMR_MiR_V3()
      $ 722 "If CMD_Unsuspend"
      if (CMD_Unsuspend):
        $ 723 "STATE≔14"
        global STATE=14
        $ 724 "ugo_update_outputs()"
        ugo_update_outputs()
      end
    elif (14 == switch_1):
      $ 725 "Case 14"
      $ 726 "Unsuspending"
      $ 727 "STATE_Info≔'Unsuspending'"
      global STATE_Info="Unsuspending"
      $ 728 "PROCESS_Step≔0"
      global PROCESS_Step=0
      $ 729 "If unsuspending()"
      if (unsuspending()):
        $ 730 "STATE≔6"
        global STATE=6
        $ 731 "ugo_update_outputs()"
        ugo_update_outputs()
      end
    elif (15 == switch_1):
      $ 732 "Case 15"
      $ 733 "Aborting"
      $ 734 "STATE_Info≔'Aborting'"
      global STATE_Info="Aborting"
      $ 735 "If aborting()"
      if (aborting()):
        $ 736 "STATE≔16"
        global STATE=16
        $ 737 "ugo_update_outputs()"
        ugo_update_outputs()
      end
    elif (16 == switch_1):
      $ 738 "Case 16"
      $ 739 "Aborted"
      $ 740 "STATE_Info≔'Aborted'"
      global STATE_Info="Aborted"
      $ 741 "If CMD_Clear"
      if (CMD_Clear):
        $ 742 "STATE≔17"
        global STATE=17
        $ 743 "ugo_update_outputs()"
        ugo_update_outputs()
      end
    elif (17 == switch_1):
      $ 744 "Case 17"
      $ 745 "Clearing"
      $ 746 "STATE_Info≔'Clearing'"
      global STATE_Info="Clearing"
      $ 747 "Clearing"
      $ 748 "reset_warning()"
      reset_warning()
      $ 749 "reset_error()"
      reset_error()
      $ 750 "If clearing()"
      if (clearing()):
        $ 751 "STATE≔2"
        global STATE=2
        $ 752 "ugo_update_outputs()"
        ugo_update_outputs()
      end
    end
    $ 753 "log_state(STATE_Info)"
    log_state(STATE_Info)
    $ 754 "log_warning(WARNING.MSG)"
    log_warning(WARNING.MSG)
    $ 755 "log_error(ERROR.MSG)"
    log_error(ERROR.MSG)
    $ 756 "Times"
    $ 757 "Switch STATE"
    switch_1 = STATE
    $ 758 "Case 1"
    if (1 == switch_1):
      $ 759 "TM_St_Stopping≔get_time(STATE_Times[STATE-1])"
      global TM_St_Stopping=get_time(STATE_Times[STATE-1])
    elif (2 == switch_1):
      $ 760 "Case 2"
      $ 761 "TM_St_Stopped≔get_time(STATE_Times[STATE-1])"
      global TM_St_Stopped=get_time(STATE_Times[STATE-1])
    elif (3 == switch_1):
      $ 762 "Case 3"
      $ 763 "TM_St_Resetting≔get_time(STATE_Times[STATE-1])"
      global TM_St_Resetting=get_time(STATE_Times[STATE-1])
    elif (4 == switch_1):
      $ 764 "Case 4"
      $ 765 "TM_St_Idle≔get_time(STATE_Times[STATE-1])"
      global TM_St_Idle=get_time(STATE_Times[STATE-1])
    elif (5 == switch_1):
      $ 766 "Case 5"
      $ 767 "TM_St_Starting≔get_time(STATE_Times[STATE-1])"
      global TM_St_Starting=get_time(STATE_Times[STATE-1])
    elif (6 == switch_1):
      $ 768 "Case 6"
      $ 769 "TM_St_Execute≔get_time(STATE_Times[STATE-1])"
      global TM_St_Execute=get_time(STATE_Times[STATE-1])
    elif (7 == switch_1):
      $ 770 "Case 7"
      $ 771 "TM_St_Completin≔get_time(STATE_Times[STATE-1])"
      global TM_St_Completin=get_time(STATE_Times[STATE-1])
    elif (8 == switch_1):
      $ 772 "Case 8"
      $ 773 "TM_St_Complete≔get_time(STATE_Times[STATE-1])"
      global TM_St_Complete=get_time(STATE_Times[STATE-1])
    elif (9 == switch_1):
      $ 774 "Case 9"
      $ 775 "TM_St_Holding≔get_time(STATE_Times[STATE-1])"
      global TM_St_Holding=get_time(STATE_Times[STATE-1])
    elif (10 == switch_1):
      $ 776 "Case 10"
      $ 777 "TM_St_Held≔get_time(STATE_Times[STATE-1])"
      global TM_St_Held=get_time(STATE_Times[STATE-1])
    elif (11 == switch_1):
      $ 778 "Case 11"
      $ 779 "TM_St_Unholding≔get_time(STATE_Times[STATE-1])"
      global TM_St_Unholding=get_time(STATE_Times[STATE-1])
    elif (12 == switch_1):
      $ 780 "Case 12"
      $ 781 "TM_St_Suspendin≔get_time(STATE_Times[STATE-1])"
      global TM_St_Suspendin=get_time(STATE_Times[STATE-1])
    elif (13 == switch_1):
      $ 782 "Case 13"
      $ 783 "TM_St_Suspended≔get_time(STATE_Times[STATE-1])"
      global TM_St_Suspended=get_time(STATE_Times[STATE-1])
    elif (14 == switch_1):
      $ 784 "Case 14"
      $ 785 "TM_St_Unsuspend≔get_time(STATE_Times[STATE-1])"
      global TM_St_Unsuspend=get_time(STATE_Times[STATE-1])
    elif (15 == switch_1):
      $ 786 "Case 15"
      $ 787 "TM_St_Aborting≔get_time(STATE_Times[STATE-1])"
      global TM_St_Aborting=get_time(STATE_Times[STATE-1])
    elif (16 == switch_1):
      $ 788 "Case 16"
      $ 789 "TM_St_Aborted≔get_time(STATE_Times[STATE-1])"
      global TM_St_Aborted=get_time(STATE_Times[STATE-1])
    elif (17 == switch_1):
      $ 790 "Case 17"
      $ 791 "TM_St_Clearing≔get_time(STATE_Times[STATE-1])"
      global TM_St_Clearing=get_time(STATE_Times[STATE-1])
    end
    $ 793 "Wait: 0.1"
    sleep(0.1)
  end
end
